Staubli VAL3: pointMove1.pgx

public program pointMove1(string x_sKey, num x_nIndex, num x_nPointIndex)
  local num l_nType
  local frame l_fFrame
  local pointRx l_pPoint
  local tool l_tTool
  local jointRx l_jJoint
  local bool l_bResult
  local jointRx l_jHere
begin
  link(l_fFrame,world)
  link(l_tTool,flange)
  //link(l_pPoint,world)
  l_nType=trajTemp:tTrajItem[x_sKey].pPointItem[x_nIndex].pParaItem.nMoveType
  call savedata:getFrame(trajTemp:tTrajItem[x_sKey].nFrameIndex,l_fFrame)
  call savedata:getTool(trajTemp:tTrajItem[x_sKey].nToolIndex,l_tTool)
  link(l_pPoint,l_fFrame)
  switch x_nPointIndex
    case 0
      l_pPoint.trsf=trajTemp:tTrajItem[x_sKey].pPointItem[x_nIndex].pInter.trsf
      l_pPoint.config=trajTemp:tTrajItem[x_sKey].pPointItem[x_nIndex].pInter.config
    break
    case 1
      l_pPoint.trsf=trajTemp:tTrajItem[x_sKey].pPointItem[x_nIndex].pPointRx.trsf
      l_pPoint.config=trajTemp:tTrajItem[x_sKey].pPointItem[x_nIndex].pPointRx.config
    break
  endSwitch

  l_jJoint=trajTemp:tTrajItem[x_sKey].pPointItem[x_nIndex].jJointRx
  if rs:_nOmacStat==9 and workingMode()==1 and isPowered()
    // if !isEmpty()
    stopMove()
    resetMotion()
    l_jHere=herej()
    movej(l_jHere,flange,mSim)
    // endIf
    //    switch l_nType
    //      case 1
    call isPointOK(x_sKey,x_nIndex,l_bResult)
    if l_bResult
      //          movel(l_pPoint,l_tTool,mSim)
      //        endIf
      //      break
      //      case 0
      movej(l_pPoint,l_tTool,mSim)
      waitEndMove()
    endIf
    //      break
    //    endSwitch
    delay(0)
  endIf
end
